FUNCTION_BLOCK TcoAbbRW_StartAtMainTask_v_8_2_x EXTENDS TcoAbbRWTask_v_8_2_x


IF Execute() THEN 
	IF _progress = 0 THEN
		IF CheckReferences() THEN
			_progress := _progress + 1;
		END_IF
	END_IF
	IF _progress = 1 THEN
		ReleaseStopCommands();
		_varInfo :=__VARINFO( inoStatus.State.AutoOn);
		THIS^.Messenger.OnCondition(_infoTimer.Q AND NOT inoStatus.State.AutoOn).Warning(_sb.Clear().Append('<#Waiting for Auto signal! #>').Append(_varInfo.Symbol).ToString());
		// Start at Main is not valid while the program is running
		_varInfo :=__VARINFO( inoStatus.State.CycleOn);
		THIS^.Messenger.OnCondition(_infoTimer.Q AND inoStatus.State.CycleOn).Warning(_sb.Clear().Append('<#Waiting for program to be stopped! #>').Append(_varInfo.Symbol).ToString());
		IF inoStatus.State.AutoOn AND NOT inoStatus.State.CycleOn THEN
			_progress := _progress + 1;
		END_IF
	END_IF
	IF _progress = 2 THEN
		IF AcquireWriteAccess() THEN
			_progress := _progress + 1;
		END_IF
	END_IF
	IF _progress = 3 THEN
		_varInfo :=__VARINFO( inoStatus.State.MotorOnState);
		THIS^.Messenger.OnCondition(_infoTimer.Q AND NOT inoStatus.State.MotorOnState).Warning(_sb.Clear().Append('<#Waiting for motors are On! #>').Append(_varInfo.Symbol).ToString());
		IF inoStatus.State.MotorOnState THEN
			_pulseTimer(IN := FALSE);
			_progress := _progress + 1;
		END_IF
	END_IF
	IF _progress = 4 THEN
		// one pulse; the controller accepts it only with write access held and the stop commands released
		inoControl.StartAtMain := Pulse();
		_varInfo :=__VARINFO( inoStatus.State.CycleOn);
		THIS^.Messenger.OnCondition(_infoTimer.Q AND NOT inoStatus.State.CycleOn).Warning(_sb.Clear().Append('<#Waiting for program running signal! #>').Append(_varInfo.Symbol).ToString());
		IF inoStatus.State.CycleOn AND NOT inoControl.StartAtMain THEN
			_progress := _progress + 1;
		END_IF
	END_IF
	IF _progress = 5 THEN
		IF ReleaseWriteAccess() THEN
			_progress := _progress + 1;
		END_IF
	END_IF

	DoneWhen(_progress = 6);
	CallTimers(TRUE);
	THIS^.ThrowWhen(_errorTimer.Q OR (_progress > 0 AND_THEN inoStatus.State.Error));
END_IF

IF  THIS^.Error AND NOT _errorMessage.Pinned THEN
	THIS^.Restore();
END_IF

METHOD PUBLIC FB_init : BOOL
VAR_INPUT
    bInitRetains : BOOL; // if TRUE, the retain variables are initialized (warm start / cold start)
    bInCopyCode : BOOL; // if TRUE, the instance afterwards gets moved into the copy code (online change)
  	ParentObject : ITcoObject;	
END_VAR
END_METHOD

(*~
	<docu>
		<summary>
			Executes when task is aborted.
		</summary>			
	</docu>	
~*)
METHOD PROTECTED OnAbort
IF  __ISVALIDREF(inoStatus) THEN   THIS^.inoStatus.ActionDescription := '<#Start at Main was aborted, while not yet completed!#>';END_IF; 
Cleanup();
END_METHOD

(*~
	<docu>
		<summary>
			Executes when task reaches the ```Done``` state .
		</summary>			
	</docu>	
~*)
METHOD PROTECTED OnDone
IF  __ISVALIDREF(inoStatus) THEN  THIS^.inoStatus.ActionDescription := '<#Start at Main was completed successfully.#>';END_IF; 
Cleanup();
_progress:=0;
END_METHOD

(*~
	<docu>
		<summary>
			Executes when task reaches the ```Error``` state.
			<para>
				Do not confuse with <see cref="PlcDocu.TcoCore.TcoTask.WhileError()"/>, that is called cyclically until '''Error''' state is left.
			</para>
		</summary>			
	</docu>	
~*)
METHOD PROTECTED OnError

VAR
	description: STRING;
END_VAR
description:= '<#Start at Main finished with error.#>';
IF  __ISVALIDREF(inoStatus) THEN   THIS^.inoStatus.ActionDescription := description; END_IF;
Cleanup();
THIS^._errorMessage.Error(_sb.Clear().Append(description).Append(' To restore acknowledge this alarm.').ToString()).Pin();
END_METHOD

METHOD PROTECTED OnStart
IF  __ISVALIDREF(inoStatus) THEN  THIS^.inoStatus.ActionDescription := '<#Start at Main started.#>'; END_IF; 
Activate();
END_METHOD

METHOD PROTECTED ReleaseCommands
inoControl.StartAtMain := FALSE;
END_METHOD

(*~
	<docu>
		<summary>
			Restores this instance to the Ready state. Can be called explicitly or from within one of the restore mechanisms.
			<para>
				See also <see cref="PlcDocu.TcoCore.TcoTask.AutoRestorable()"/>
			</para>
		</summary>			
	</docu>	
~*)
METHOD Restore : ITcoRestorable
SUPER^.Restore();
END_METHOD

END_FUNCTION_BLOCK

(* stored: Version 1.1.0.1, ProductVersion 3.1.4024.12
   POU TcoAbbRW_StartAtMainTask_v_8_2_x: Id {5386d75b-229e-4d90-a779-599a9cc8e842}, SpecialFunc None
   Method FB_init: Id {47f18b16-c760-416d-9945-93f5a2be79a7}
   Method OnAbort: Id {7012e2db-d11d-4c39-8fcf-4ab81b2ec35d}
   Method OnDone: Id {8c677c2d-8657-4ab5-bd14-883024544c7b}
   Method OnError: Id {6ef1232b-51a3-44fe-9fe6-f85e2d0d3d44}
   Method OnStart: Id {50a9481d-163a-4c09-8a1f-a67d311d4ccf}
   Method ReleaseCommands: Id {47221457-0da7-4050-b7e2-c7c270da56b1}
   Method Restore: Id {03126fac-693a-48f3-853b-bfff768debae} *)
